DATA_BLOCK "naut_Tags"
{ S7_Optimized_Access := 'TRUE' }
VERSION : 0.1
   VAR
      Reset : BOOL;
      Running : BOOL;
      Start : BOOL;
   END_VAR

BEGIN

END_DATA_BLOCK
